// TIA Portal V20 export
ORGANIZATION_BLOCK "T10_Ciclo"   // OB131, LAD, ProgramCycle
TITLE = T10_Ciclo
{ S7_Optimized_Access := 'TRUE' }
AUTHOR : IA
FAMILY : PRUEBA
VERSION : 0.1
// Tanda 4B: comunicación del PLC consigo mismo
// stored: AutoNumber false, IsIECCheckEnabled false, SetENOAutomatically false
   VAR_INPUT
      Initial_Call : Bool;
      Remanence : Bool;
   END_VAR
BEGIN

REGION Network 1: T10_Llamar
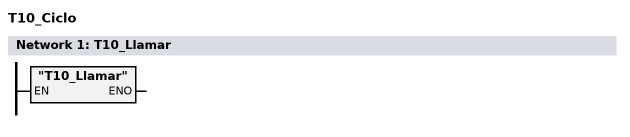
   RUNG wire#powerrail
      "T10_Llamar"()
   END_RUNG
   // the same network as SCL:
   "T10_Llamar"();
END_REGION
END_ORGANIZATION_BLOCK
